// TIA Portal V21 export
// export: Created 2026-08-21T20:18:50.5747954Z, ExportSetting None, DisplayName Totally Integrated Automation Portal, DisplayVersion V21, DisplayName STEP 7 Professional, DisplayVersion V21, DisplayName STEP 7 Safety, DisplayVersion V21, DisplayName Tech WebApplication, DisplayVersion V21, DisplayName WinCC Basic/Comfort/Advanced, DisplayVersion V21, DisplayName WinCC Professional, DisplayVersion V21, DisplayName WinCC Unified, DisplayVersion V21
FUNCTION "ConvertToStruCm" : Void   // FC20, SCL
{ S7_Optimized_Access := 'TRUE' }
// stored: SetENOAutomatically false
   VAR_INPUT
      AnaVal1 : "AnaVal";   // Rbk
      AnaVal2 : "AnaVal";
      AnaVal3 : "AnaVal";
      DigVal1 : "DigVal";
      DigVal2 : "DigVal";
      DigVal3 : "DigVal";
      Scale : "ScaVal";   // MV_Scale
      ScaleRAW : "ScaVal_Raw";   // MV_ScaleRAW
      Unit : Int;   // MV_Unit
   END_VAR
   VAR_OUTPUT
      StruCm_Out : "StruCm";
   END_VAR
BEGIN
   #StruCm_Out.AnaVal1 := #AnaVal1;
   #StruCm_Out.AnaVal2 := #AnaVal2;
   #StruCm_Out.AnaVal3 := #AnaVal3;
   #StruCm_Out.DigVal1 := #DigVal1;
   #StruCm_Out.DigVal2 := #DigVal2;
   #StruCm_Out.DigVal3 := #DigVal3;
   #StruCm_Out.Scale := #Scale;
   #StruCm_Out.ScaleRAW := #ScaleRAW;
   #StruCm_Out.Unit := #Unit;
END_FUNCTION
